FUNCTION_BLOCK STAR_DELTA (* Migrated from IEC 61131-3 ST *)
  (* Standard: 61499-2 *)
  (* Version 1.0, 2026-11-06, st2fb *)
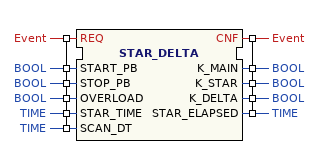
  EVENT_INPUT
    REQ WITH START_PB, STOP_PB, OVERLOAD, STAR_TIME, SCAN_DT;
  END_EVENT
  EVENT_OUTPUT
    CNF WITH K_MAIN, K_STAR, K_DELTA, STAR_ELAPSED;
  END_EVENT
  VAR_INPUT
    START_PB : BOOL;
    STOP_PB : BOOL;
    OVERLOAD : BOOL;
    STAR_TIME : TIME;
    SCAN_DT : TIME;
  END_VAR
  VAR_OUTPUT
    K_MAIN : BOOL;
    K_STAR : BOOL;
    K_DELTA : BOOL;
    STAR_ELAPSED : TIME;
  END_VAR
  VAR
    RUN_CMD : BOOL := FALSE;
    ST2FB_NOW : TIME := T#0s;
    STAR_TIMER_IN : BOOL := FALSE;
    STAR_TIMER_PT : TIME := T#0s;
    STAR_TIMER_Q : BOOL := FALSE;
    STAR_TIMER_ET : TIME := T#0s;
    STAR_TIMER_STATE : INT := 0;
    STAR_TIMER_PREV_IN : BOOL := FALSE;
    STAR_TIMER_START_TIME : TIME := T#0s;
    GAP_TIMER_IN : BOOL := FALSE;
    GAP_TIMER_PT : TIME := T#0s;
    GAP_TIMER_Q : BOOL := FALSE;
    GAP_TIMER_ET : TIME := T#0s;
    GAP_TIMER_STATE : INT := 0;
    GAP_TIMER_PREV_IN : BOOL := FALSE;
    GAP_TIMER_START_TIME : TIME := T#0s;
  END_VAR
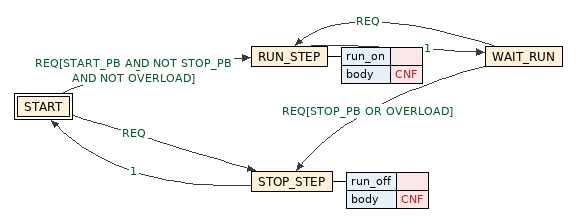
  EC_STATES
    START;
    RUN_STEP : run_on, body -> CNF;
    WAIT_RUN;
    STOP_STEP : run_off, body -> CNF;
  END_STATES
  EC_TRANSITIONS
    START TO RUN_STEP := REQ[START_PB AND NOT STOP_PB AND NOT OVERLOAD];
    START TO STOP_STEP := REQ;
    RUN_STEP TO WAIT_RUN := 1;
    WAIT_RUN TO STOP_STEP := REQ[STOP_PB OR OVERLOAD];
    WAIT_RUN TO RUN_STEP := REQ;
    STOP_STEP TO START := 1;
  END_TRANSITIONS
  ALGORITHM run_on IN ST:
ST2FB_NOW := ST2FB_NOW + SCAN_DT;
RUN_CMD := TRUE;
  END_ALGORITHM
  ALGORITHM run_off IN ST:
ST2FB_NOW := ST2FB_NOW + SCAN_DT;
RUN_CMD := FALSE;
  END_ALGORITHM
  ALGORITHM body IN ST:
STAR_TIMER_IN := RUN_CMD;
STAR_TIMER_PT := STAR_TIME;
IF (STAR_TIMER_STATE = 0) AND NOT STAR_TIMER_PREV_IN AND STAR_TIMER_IN THEN
  STAR_TIMER_STATE := 1;
  STAR_TIMER_Q := FALSE;
  STAR_TIMER_START_TIME := ST2FB_NOW;
ELSE
  IF NOT STAR_TIMER_IN THEN
    STAR_TIMER_ET := T#0s;
    STAR_TIMER_Q := FALSE;
    STAR_TIMER_STATE := 0;
  ELSIF STAR_TIMER_STATE = 1 THEN
    IF STAR_TIMER_START_TIME + STAR_TIMER_PT <= ST2FB_NOW THEN
      STAR_TIMER_STATE := 2;
      STAR_TIMER_Q := TRUE;
      STAR_TIMER_ET := STAR_TIMER_PT;
    ELSE
      STAR_TIMER_ET := ST2FB_NOW - STAR_TIMER_START_TIME;
    END_IF;
  END_IF;
END_IF;
STAR_TIMER_PREV_IN := STAR_TIMER_IN;
GAP_TIMER_IN := STAR_TIMER_Q;
GAP_TIMER_PT := T#50ms;
IF (GAP_TIMER_STATE = 0) AND NOT GAP_TIMER_PREV_IN AND GAP_TIMER_IN THEN
  GAP_TIMER_STATE := 1;
  GAP_TIMER_Q := FALSE;
  GAP_TIMER_START_TIME := ST2FB_NOW;
ELSE
  IF NOT GAP_TIMER_IN THEN
    GAP_TIMER_ET := T#0s;
    GAP_TIMER_Q := FALSE;
    GAP_TIMER_STATE := 0;
  ELSIF GAP_TIMER_STATE = 1 THEN
    IF GAP_TIMER_START_TIME + GAP_TIMER_PT <= ST2FB_NOW THEN
      GAP_TIMER_STATE := 2;
      GAP_TIMER_Q := TRUE;
      GAP_TIMER_ET := GAP_TIMER_PT;
    ELSE
      GAP_TIMER_ET := ST2FB_NOW - GAP_TIMER_START_TIME;
    END_IF;
  END_IF;
END_IF;
GAP_TIMER_PREV_IN := GAP_TIMER_IN;
K_MAIN := RUN_CMD;
K_STAR := RUN_CMD AND NOT STAR_TIMER_Q;
K_DELTA := RUN_CMD AND GAP_TIMER_Q;
STAR_ELAPSED := STAR_TIMER_ET;
  END_ALGORITHM
END_FUNCTION_BLOCK
